Fanuc KAREL source: kt00005.KL

-- PROVISIONAL review KL for V770-1; original PC SHA256 3043a2a622869e48eea76a28951aaa6a1838e524b5c196e3bcbe4c44e792f88d
-- Incomplete behavior may be omitted. Consult companion uncertainty JSON. Do not deploy.
PROGRAM KT00005
%NOLOCKGROUP
VAR
  I1 : INTEGER
  OUT : INTEGER
-- UNRESOLVED_DECL Y2 type=002018
BEGIN
  -- UNRESOLVED_PC offsets 5-16; opcodes 2E,23
  -- UNRESOLVED_PC offsets 21-35; opcodes 2E,22,9D,33,B2
  -- UNRESOLVED_PC offsets 40-62; opcodes 21,22,9D,33,B1,52,23
  -- UNRESOLVED_PC offsets 67-71; opcodes 7F
END KT00005
